PROGRAM main
  VAR
    S1 AT %IX0.0 : BOOL; (* pulsador NA *)
    H1 AT %QX0.0 : BOOL; (* luz que cambia al apretar *)
    H2 AT %QX0.1 : BOOL; (* luz que cambia al soltar *)
    APRIETA      : R_TRIG;
    SUELTA       : F_TRIG;
    PULSO        : BOOL; (* un ciclo al apretar *)
    PULSO2       : BOOL; (* un ciclo al soltar *)
  END_VAR
  VAR  (* added by the conversion: wires and edge detectors of the diagram *)
    R_TRIG1 : R_TRIG;
  END_VAR

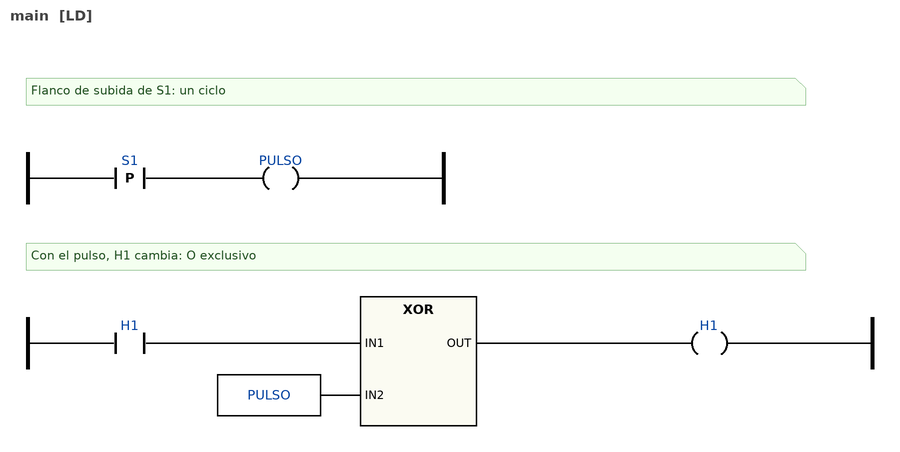
(* LD diagram, written out as Structured Text *)
(* Flanco de subida de S1: un ciclo *)
R_TRIG1(CLK := S1);
PULSO := R_TRIG1.Q;
(* Con el pulso, H1 cambia: O exclusivo *)
H1 := H1 XOR PULSO;
END_PROGRAM
